(* IEC 61131-3 sources: codesys-to-s7/tests/corpus/C2S7-POU-STAT/neg, 1 file *)

(* ---- input.st ---- *)
FUNCTION_BLOCK FB_Case
VAR
    n : INT;
END_VAR
n := n + 1;
END_FUNCTION_BLOCK
